TEXTLIST TextList_StateLong_1
  0 = 'Not Clean'
  7 = 'Clean'
  9 = 'Product'
   = ''
END_TEXTLIST

(* stored: Version 1.1.0.1, ProductVersion 3.1.4024.12
   TextList TextList_StateLong_1: Id {a0610e6c-4e8a-47ff-8adf-a29587a18e06} *)
